// TIA Portal V20 export
DATA_BLOCK "T2_Resultado"   // DB40923
{ S7_Optimized_Access := 'TRUE' }
AUTHOR : IA
FAMILY : PRUEBA
VERSION : 0.1
// Prueba IA 2: un Bool por prueba. Base_Todo_OK = todo correcto
// stored: AutoNumber false
   VAR
      T01_Contacto : Bool;   // Contacto NA con TRUE
      T02_Contacto_negado : Bool;   // Contacto NC sobre bit FALSE
      T03_Not : Bool;   // Inversor NOT
      T04_Set : Bool;   // Bobina S (set)
      T05_Reset : Bool;   // Bobina R (reset)
      T06_Flanco_P : Bool;   // Flanco positivo PBox (un ciclo, enclavado)
      T07_Serie_AND : Bool;   // Dos contactos en serie
      T08_Variable_PLC : Bool;   // Variable %M de la tabla T2_Variables
      T09_Eq_Int : Bool;   // Igual (Int)
      T10_Ne_Word : Bool;   // Distinto (Word)
      T11_Gt_Real : Bool;   // Mayor (Real)
      T12_Ge_DInt : Bool;   // Mayor o igual (DInt)
      T13_Lt_Int : Bool;   // Menor (Int)
      T14_Rango : Bool;   // Dos comparaciones en serie (rango)
      T15_Move : Bool;   // Move (1 salida)
      T16_Move_2_salidas : Bool;   // Move (2 salidas)
      T17_Swap : Bool;   // Swap de bytes (Word)
      T18_Convert : Bool;   // Convert Int -> Real
      T19_S_Move_LEN : Bool;   // S_Move de String y LEN
      T20_Serialize_Deserialize : Bool;   // Serialize + Deserialize de un UDT anidado
      T21_Calculate : Bool;   // Calculate (IN1*IN2)+IN3
      T22_Add : Bool;   // Suma (Add)
      T23_Sub : Bool;   // Resta (Sub)
      T24_CONCAT : Bool;   // CONCAT de dos String
      T25_VAL_STRG_STRG_VAL : Bool;   // Número -> texto -> número
      T26_MAX_LEN : Bool;   // MAX_LEN de String[20]
      T27_Strg_TO_Chars : Bool;   // String -> Array of Char
      T28_TON : Bool;   // TON (IEC_TIMER en DB global)
      T29_RD_SYS_T : Bool;   // Leer hora del sistema (DTL)
      T30_Llamada_FC : Bool;   // Llamada a FC SCL con parámetros
      T31_Llamada_FB_KOP : Bool;   // FB KOP (SD) con DB de instancia (SD) y TON interno
      T32_Llamada_FB_SCL : Bool;   // FB SCL (fuente) con DB de instancia
      T33_SCL_IF : Bool;   // SCL: IF / ELSIF / ELSE
      T34_SCL_CASE : Bool;   // SCL: CASE
      T35_SCL_FOR_WHILE : Bool;   // SCL: FOR y WHILE
      T36_SCL_String : Bool;   // SCL: CONCAT, LEN, LEFT
      T37_SCL_Real : Bool;   // SCL: SQRT y operaciones Real
      T38_SCL_Slice : Bool;   // SCL: acceso a bit %X de un Word
      T39_SCL_Funcion : Bool;   // SCL: llamada a FC con valor de retorno
      T40_SCL_Array_UDT : Bool;   // SCL: array de UDT
      T41_SCL_Conversion : Bool;   // SCL: conversiones de tipo
      N01_OR_ramas : Bool;   // [NUEVA] OR con dos ramas en paralelo
      N02_Mul : Bool;   // [NUEVA] Multiplicación (Mul)
      N03_Div : Bool;   // [NUEVA] División (Div)
      N04_Le : Bool;   // [NUEVA] Menor o igual (Le)
      N05_FC_retorno_KOP : Bool;   // [NUEVA] Llamada KOP a FC con valor de retorno
      Base_OK : Int;   // Pruebas base correctas
      Base_Total : Int := 41;   // Pruebas base
      Base_Todo_OK : Bool;   // TRUE si todas las base están bien
      Nuevas_OK : Int;   // Pruebas nuevas correctas
      Nuevas_Total : Int := 5;   // Pruebas nuevas
      Vida_OB125 : DInt;   // Sube 1 en cada ciclo si el OB125 se ejecuta
      Vida_T2_Bits : DInt;   // Sube 1 en cada ciclo si T2_Bits se ejecuta
   END_VAR
BEGIN
END_DATA_BLOCK
